(* IEC 61131-3 sources: plc-st-coding-agent/progress/evidence/f14_v13_self_20261113/jobs/custom_deepseek-v4pro (part 2) *)

(* ---- public-hard-01.raw_candidate_02.st ---- *)
(*
ENGINEERING_CONTRACT
Outputs/state group | activation | retention/hold | reset/deactivation | same-scan priority | units/bounds
estop: highest priority; active-low; all outputs false and internal states/latches reset (PUB001, PUB003).
Manual valve/motor: rising button toggles local latch; held between scans; reset by estop or mode change (PUB002, PUB004-PUB005).
AutoState: idle all off; fillA A on until level>=50; fillB B on until level>=80; processMode false->mix, true->fillC C on until level>=100; mix motor on until complete signal false->true while motor running; deliver D on and retained until autoStart/estop/mode change (PUB006-PUB015).
AutoStart rising restarts at fillA and suppresses threshold transition for first scan; transitions update state before output mapping this scan.
levelSensor INT cm; thresholds use >=.
mix completion uses armed condition requiring mixMotorComplete FALSE before TRUE while in mix state.
*)
(* CONTRACT_RULES [] *)
FUNCTION_BLOCK MaterialProportioningControl
VAR_INPUT
    estop : BOOL;
    opeMode : BOOL;
    valveAStart : BOOL;
    valveBStart : BOOL;
    valveCStart : BOOL;
    valveDStart : BOOL;
    mixMotorStart : BOOL;
    autoStart : BOOL;
    processMode : BOOL;
    levelSensor : INT;
    mixMotorComplete : BOOL;
END_VAR
VAR_OUTPUT
    valveARun : BOOL;
    valveBRun : BOOL;
    valveCRun : BOOL;
    valveDRun : BOOL;
    mixMotorRun : BOOL;
END_VAR
VAR CONSTANT
    AUTO_IDLE : INT := 0;
    AUTO_FILL_A : INT := 1;
    AUTO_FILL_B : INT := 2;
    AUTO_FILL_C : INT := 3;
    AUTO_MIX : INT := 4;
    AUTO_DELIVER : INT := 5;
END_VAR
VAR
    autoStartRtr : R_TRIG;
    valveAStartRtr : R_TRIG;
    valveBStartRtr : R_TRIG;
    valveCStartRtr : R_TRIG;
    valveDStartRtr : R_TRIG;
    mixMotorStartRtr : R_TRIG;

    local_prevOpeMode : BOOL := FALSE;
    local_init : BOOL := FALSE;

    local_manualA : BOOL := FALSE;
    local_manualB : BOOL := FALSE;
    local_manualC : BOOL := FALSE;
    local_manualD : BOOL := FALSE;
    local_manualMix : BOOL := FALSE;

    local_autoState : INT := AUTO_IDLE;
    local_firstAutoScan : BOOL := FALSE;
    local_mixArmed : BOOL := FALSE;

    local_autoStartEdge : BOOL;
    local_edgeA : BOOL;
    local_edgeB : BOOL;
    local_edgeC : BOOL;
    local_edgeD : BOOL;
    local_edgeMix : BOOL;
END_VAR

autoStartRtr(CLK := autoStart);
valveAStartRtr(CLK := valveAStart);
valveBStartRtr(CLK := valveBStart);
valveCStartRtr(CLK := valveCStart);
valveDStartRtr(CLK := valveDStart);
mixMotorStartRtr(CLK := mixMotorStart);

local_autoStartEdge := autoStartRtr.Q AND opeMode AND estop;
local_edgeA := valveAStartRtr.Q AND NOT opeMode AND estop;
local_edgeB := valveBStartRtr.Q AND NOT opeMode AND estop;
local_edgeC := valveCStartRtr.Q AND NOT opeMode AND estop;
local_edgeD := valveDStartRtr.Q AND NOT opeMode AND estop;
local_edgeMix := mixMotorStartRtr.Q AND NOT opeMode AND estop;

IF NOT local_init THEN
    local_prevOpeMode := opeMode;
    local_init := TRUE;
ELSIF local_prevOpeMode <> opeMode THEN
    local_prevOpeMode := opeMode;
    local_manualA := FALSE;
    local_manualB := FALSE;
    local_manualC := FALSE;
    local_manualD := FALSE;
    local_manualMix := FALSE;
    local_autoState := AUTO_IDLE;
    local_firstAutoScan := FALSE;
    local_mixArmed := FALSE;
END_IF;

IF NOT estop THEN
    valveARun := FALSE;
    valveBRun := FALSE;
    valveCRun := FALSE;
    valveDRun := FALSE;
    mixMotorRun := FALSE;

    local_manualA := FALSE;
    local_manualB := FALSE;
    local_manualC := FALSE;
    local_manualD := FALSE;
    local_manualMix := FALSE;
    local_autoState := AUTO_IDLE;
    local_firstAutoScan := FALSE;
    local_mixArmed := FALSE;
    RETURN;
END_IF;

IF opeMode THEN
    IF local_autoStartEdge THEN
        local_autoState := AUTO_FILL_A;
        local_firstAutoScan := TRUE;
        local_mixArmed := FALSE;
    END_IF;

    IF NOT local_firstAutoScan THEN
        IF local_autoState = AUTO_FILL_A THEN
            IF levelSensor >= 50 THEN
                local_autoState := AUTO_FILL_B;
            END_IF;
        ELSIF local_autoState = AUTO_FILL_B THEN
            IF levelSensor >= 80 THEN
                IF processMode THEN
                    local_autoState := AUTO_FILL_C;
                ELSE
                    local_autoState := AUTO_MIX;
                END_IF;
            END_IF;
        ELSIF local_autoState = AUTO_FILL_C THEN
            IF levelSensor >= 100 THEN
                local_autoState := AUTO_MIX;
            END_IF;
        ELSIF local_autoState = AUTO_MIX THEN
            IF local_mixArmed AND mixMotorComplete THEN
                local_autoState := AUTO_DELIVER;
            END_IF;
        END_IF;
    END_IF;

    IF local_autoState = AUTO_MIX THEN
        IF NOT mixMotorComplete THEN
            local_mixArmed := TRUE;
        END_IF;
    ELSE
        local_mixArmed := FALSE;
    END_IF;

    CASE local_autoState OF
        AUTO_IDLE:
            valveARun := FALSE;
            valveBRun := FALSE;
            valveCRun := FALSE;
            valveDRun := FALSE;
            mixMotorRun := FALSE;

        AUTO_FILL_A:
            valveARun := TRUE;
            valveBRun := FALSE;
            valveCRun := FALSE;
            valveDRun := FALSE;
            mixMotorRun := FALSE;

        AUTO_FILL_B:
            valveARun := FALSE;
            valveBRun := TRUE;
            valveCRun := FALSE;
            valveDRun := FALSE;
            mixMotorRun := FALSE;

        AUTO_FILL_C:
            valveARun := FALSE;
            valveBRun := FALSE;
            valveCRun := TRUE;
            valveDRun := FALSE;
            mixMotorRun := FALSE;

        AUTO_MIX:
            valveARun := FALSE;
            valveBRun := FALSE;
            valveCRun := FALSE;
            valveDRun := FALSE;
            mixMotorRun := TRUE;

        AUTO_DELIVER:
            valveARun := FALSE;
            valveBRun := FALSE;
            valveCRun := FALSE;
            valveDRun := TRUE;
            mixMotorRun := FALSE;
    END_CASE;

    local_firstAutoScan := FALSE;
ELSE
    IF local_edgeA THEN
        local_manualA := NOT local_manualA;
    END_IF;

    IF local_edgeB THEN
        local_manualB := NOT local_manualB;
    END_IF;

    IF local_edgeC THEN
        local_manualC := NOT local_manualC;
    END_IF;

    IF local_edgeD THEN
        local_manualD := NOT local_manualD;
    END_IF;

    IF local_edgeMix THEN
        local_manualMix := NOT local_manualMix;
    END_IF;

    valveARun := local_manualA;
    valveBRun := local_manualB;
    valveCRun := local_manualC;
    valveDRun := local_manualD;
    mixMotorRun := local_manualMix;
END_IF;
END_FUNCTION_BLOCK

(* ---- public-hard-02.candidate_01.st ---- *)
(*
ENGINEERING_CONTRACT
- State machine: 0=IDLE, 1=MOVING, 2=WAIT_COMPLETE, 3=DONE.
- IDLE->MOVING on rising edge of station1Start while sensor1; loads first active entry (PUB001).
- MOVING drives conveyor direction from targetStation-currentStation; stops same scan target sensor TRUE (PUB002/PUB005).
- Arrival at stations 2..4 enters WAIT_COMPLETE; arrival at 5 enters DONE (PUB003).
- WAIT_COMPLETE waits for the matching stationXComplete rising edge, then loads next entry; final 5 ends DONE (PUB003).
- Conveyor outputs are state/direction combinational and are not retained once movement stops; opposite directions cannot overlap (PUB004, V12.1).
- No unstated reset or new-cycle restart after DONE.
- Inputs are assumed valid: processLength 1..8, entries 2..5, final 5.
*)
(* CONTRACT_RULES [] *)
FUNCTION_BLOCK FlexibleProcessingControl
VAR_INPUT
    processLength : USINT;
    sensor1 : BOOL;
    sensor2 : BOOL;
    sensor3 : BOOL;
    sensor4 : BOOL;
    sensor5 : BOOL;
    station1Start : BOOL;
    station2Complete : BOOL;
    station3Complete : BOOL;
    station4Complete : BOOL;
    processSequence : ARRAY[1..8] OF USINT;
END_VAR
VAR_OUTPUT
    conveyorLeft : BOOL;
    conveyorRight : BOOL;
END_VAR
VAR
    state : INT := 0; (* 0 IDLE, 1 MOVING, 2 WAIT_COMPLETE, 3 DONE *)
    idx : USINT := 1;
    currentStation : USINT := 1;
    targetStation : USINT := 5;
    directionRight : BOOL := TRUE;
    targetArrived : BOOL := FALSE;
    completionQ : BOOL := FALSE;
    startTrig : R_TRIG;
    comp2Trig : R_TRIG;
    comp3Trig : R_TRIG;
    comp4Trig : R_TRIG;
END_VAR

startTrig(CLK := station1Start);
comp2Trig(CLK := station2Complete);
comp3Trig(CLK := station3Complete);
comp4Trig(CLK := station4Complete);

CASE targetStation OF
    2: targetArrived := sensor2;
    3: targetArrived := sensor3;
    4: targetArrived := sensor4;
    5: targetArrived := sensor5;
ELSE
    targetArrived := FALSE;
END_CASE;

IF processLength = 0 OR processLength > 8 THEN
    state := 3;
ELSE
    CASE state OF
        0: (* IDLE *)
            IF startTrig.Q AND sensor1 THEN
                idx := 1;
                currentStation := 1;
                targetStation := processSequence[idx];
                IF targetStation >= 2 AND targetStation <= 5 THEN
                    directionRight := targetStation > currentStation;
                    CASE targetStation OF
                        2: targetArrived := sensor2;
                        3: targetArrived := sensor3;
                        4: targetArrived := sensor4;
                        5: targetArrived := sensor5;
                    END_CASE;
                    IF targetArrived THEN
                        currentStation := targetStation;
                        IF targetStation = 5 THEN
                            state := 3;
                        ELSE
                            state := 2;
                        END_IF;
                    ELSE
                        state := 1;
                    END_IF;
                ELSE
                    state := 3;
                END_IF;
            END_IF;

        1: (* MOVING *)
            IF targetArrived THEN
                currentStation := targetStation;
                IF targetStation = 5 THEN
                    state := 3;
                ELSE
                    state := 2;
                END_IF;
            END_IF;

        2: (* WAIT_COMPLETE *)
            completionQ := FALSE;
            CASE currentStation OF
                2: completionQ := comp2Trig.Q;
                3: completionQ := comp3Trig.Q;
                4: completionQ := comp4Trig.Q;
            ELSE
                state := 3;
            END_CASE;
            IF completionQ THEN
                idx := idx + 1;
                IF idx > processLength THEN
                    state := 3;
                ELSE
                    targetStation := processSequence[idx];
                    IF targetStation >= 2 AND targetStation <= 5 THEN
                        directionRight := targetStation > currentStation;
                        CASE targetStation OF
                            2: targetArrived := sensor2;
                            3: targetArrived := sensor3;
                            4: targetArrived := sensor4;
                            5: targetArrived := sensor5;
                        END_CASE;
                        IF targetArrived THEN
                            currentStation := targetStation;
                            IF targetStation = 5 THEN
                                state := 3;
                            ELSE
                                state := 2;
                            END_IF;
                        ELSE
                            state := 1;
                        END_IF;
                    ELSE
                        state := 3;
                    END_IF;
                END_IF;
            END_IF;

        3: (* DONE *)
            (* no action *)
    END_CASE;
END_IF;

IF state = 1 THEN
    IF directionRight THEN
        conveyorRight := TRUE;
        conveyorLeft := FALSE;
    ELSE
        conveyorLeft := TRUE;
        conveyorRight := FALSE;
    END_IF;
ELSE
    conveyorLeft := FALSE;
    conveyorRight := FALSE;
END_IF;

END_FUNCTION_BLOCK

(* ---- public-hard-02.candidate_03.st ---- *)
(*
ENGINEERING_CONTRACT
- State machine: 0=IDLE, 1=MOVING, 2=WAIT_COMPLETE, 3=DONE.
- IDLE->MOVING on rising edge of station1Start while sensor1; loads first active entry (PUB001).
- MOVING drives conveyor direction from targetStation-currentStation; stops same scan target sensor TRUE (PUB002/PUB005).
- Arrival at stations 2..4 enters WAIT_COMPLETE; arrival at 5 enters DONE (PUB003).
- WAIT_COMPLETE waits for the matching stationXComplete rising edge, then loads next entry; final 5 ends DONE (PUB003).
- Conveyor outputs are state/direction combinational and are not retained once movement stops; opposite directions cannot overlap (PUB004, V12.1).
- No unstated reset or new-cycle restart after DONE.
- Inputs are assumed valid: processLength 1..8, entries 2..5, final 5.
*)
(* CONTRACT_RULES [] *)
FUNCTION_BLOCK FlexibleProcessingControl
VAR_INPUT
    processLength : USINT;
    sensor1 : BOOL;
    sensor2 : BOOL;
    sensor3 : BOOL;
    sensor4 : BOOL;
    sensor5 : BOOL;
    station1Start : BOOL;
    station2Complete : BOOL;
    station3Complete : BOOL;
    station4Complete : BOOL;
    processSequence : ARRAY[1..8] OF USINT;
END_VAR
VAR_OUTPUT
    conveyorLeft : BOOL;
    conveyorRight : BOOL;
END_VAR
VAR
    state : INT := 0; (* 0 IDLE, 1 MOVING, 2 WAIT_COMPLETE, 3 DONE *)
    idx : USINT := 1;
    currentStation : USINT := 1;
    targetStation : USINT := 5;
    directionRight : BOOL := TRUE;
    targetArrived : BOOL := FALSE;
    completionQ : BOOL := FALSE;
    startTrig : R_TRIG;
    comp2Trig : R_TRIG;
    comp3Trig : R_TRIG;
    comp4Trig : R_TRIG;
END_VAR

startTrig(CLK := station1Start);
comp2Trig(CLK := station2Complete);
comp3Trig(CLK := station3Complete);
comp4Trig(CLK := station4Complete);

CASE targetStation OF
    2: targetArrived := sensor2;
    3: targetArrived := sensor3;
    4: targetArrived := sensor4;
    5: targetArrived := sensor5;
ELSE
    targetArrived := FALSE;
END_CASE;

IF processLength = 0 OR processLength > 8 THEN
    state := 3;
ELSE
    CASE state OF
        0: (* IDLE *)
            IF startTrig.Q AND sensor1 THEN
                idx := 1;
                currentStation := 1;
                targetStation := processSequence[idx];
                IF targetStation >= 2 AND targetStation <= 5 THEN
                    directionRight := targetStation > currentStation;
                    CASE targetStation OF
                        2: targetArrived := sensor2;
                        3: targetArrived := sensor3;
                        4: targetArrived := sensor4;
                        5: targetArrived := sensor5;
                    END_CASE;
                    IF targetArrived THEN
                        currentStation := targetStation;
                        IF targetStation = 5 THEN
                            state := 3;
                        ELSE
                            state := 2;
                        END_IF;
                    ELSE
                        state := 1;
                    END_IF;
                ELSE
                    state := 3;
                END_IF;
            END_IF;

        1: (* MOVING *)
            IF targetArrived THEN
                currentStation := targetStation;
                IF targetStation = 5 THEN
                    state := 3;
                ELSE
                    state := 2;
                END_IF;
            END_IF;

        2: (* WAIT_COMPLETE *)
            completionQ := FALSE;
            CASE currentStation OF
                2: completionQ := comp2Trig.Q;
                3: completionQ := comp3Trig.Q;
                4: completionQ := comp4Trig.Q;
            ELSE
                state := 3;
            END_CASE;
            IF completionQ THEN
                idx := idx + 1;
                IF idx > processLength THEN
                    state := 3;
                ELSE
                    targetStation := processSequence[idx];
                    IF targetStation >= 2 AND targetStation <= 5 THEN
                        IF targetStation = currentStation THEN
                            targetArrived := TRUE;
                        ELSE
                            directionRight := targetStation > currentStation;
                            CASE targetStation OF
                                2: targetArrived := sensor2;
                                3: targetArrived := sensor3;
                                4: targetArrived := sensor4;
                                5: targetArrived := sensor5;
                            END_CASE;
                        END_IF;
                        IF targetArrived THEN
                            currentStation := targetStation;
                            IF targetStation = 5 THEN
                                state := 3;
                            ELSE
                                state := 2;
                            END_IF;
                        ELSE
                            state := 1;
                        END_IF;
                    ELSE
                        state := 3;
                    END_IF;
                END_IF;
            END_IF;

        3: (* DONE *)
            state := 0;
    END_CASE;
END_IF;

IF state = 1 THEN
    IF directionRight THEN
        conveyorRight := TRUE;
        conveyorLeft := FALSE;
    ELSE
        conveyorLeft := TRUE;
        conveyorRight := FALSE;
    END_IF;
ELSE
    conveyorLeft := FALSE;
    conveyorRight := FALSE;
END_IF;

END_FUNCTION_BLOCK

(* ---- public-hard-02.patch_base_02.st ---- *)
(*
ENGINEERING_CONTRACT
- State machine: 0=IDLE, 1=MOVING, 2=WAIT_COMPLETE, 3=DONE.
- IDLE->MOVING on rising edge of station1Start while sensor1; loads first active entry (PUB001).
- MOVING drives conveyor direction from targetStation-currentStation; stops same scan target sensor TRUE (PUB002/PUB005).
- Arrival at stations 2..4 enters WAIT_COMPLETE; arrival at 5 enters DONE (PUB003).
- WAIT_COMPLETE waits for the matching stationXComplete rising edge, then loads next entry; final 5 ends DONE (PUB003).
- Conveyor outputs are state/direction combinational and are not retained once movement stops; opposite directions cannot overlap (PUB004, V12.1).
- No unstated reset or new-cycle restart after DONE.
- Inputs are assumed valid: processLength 1..8, entries 2..5, final 5.
*)
(* CONTRACT_RULES [] *)
FUNCTION_BLOCK FlexibleProcessingControl
VAR_INPUT
    processLength : USINT;
    sensor1 : BOOL;
    sensor2 : BOOL;
    sensor3 : BOOL;
    sensor4 : BOOL;
    sensor5 : BOOL;
    station1Start : BOOL;
    station2Complete : BOOL;
    station3Complete : BOOL;
    station4Complete : BOOL;
    processSequence : ARRAY[1..8] OF USINT;
END_VAR
VAR_OUTPUT
    conveyorLeft : BOOL;
    conveyorRight : BOOL;
END_VAR
VAR
    state : INT := 0; (* 0 IDLE, 1 MOVING, 2 WAIT_COMPLETE, 3 DONE *)
    idx : USINT := 1;
    currentStation : USINT := 1;
    targetStation : USINT := 5;
    directionRight : BOOL := TRUE;
    targetArrived : BOOL := FALSE;
    completionQ : BOOL := FALSE;
    startTrig : R_TRIG;
    comp2Trig : R_TRIG;
    comp3Trig : R_TRIG;
    comp4Trig : R_TRIG;
END_VAR

startTrig(CLK := station1Start);
comp2Trig(CLK := station2Complete);
comp3Trig(CLK := station3Complete);
comp4Trig(CLK := station4Complete);

CASE targetStation OF
    2: targetArrived := sensor2;
    3: targetArrived := sensor3;
    4: targetArrived := sensor4;
    5: targetArrived := sensor5;
ELSE
    targetArrived := FALSE;
END_CASE;

IF processLength = 0 OR processLength > 8 THEN
    state := 3;
ELSE
    CASE state OF
        0: (* IDLE *)
            IF startTrig.Q AND sensor1 THEN
                idx := 1;
                currentStation := 1;
                targetStation := processSequence[idx];
                IF targetStation >= 2 AND targetStation <= 5 THEN
                    directionRight := targetStation > currentStation;
                    CASE targetStation OF
                        2: targetArrived := sensor2;
                        3: targetArrived := sensor3;
                        4: targetArrived := sensor4;
                        5: targetArrived := sensor5;
                    END_CASE;
                    IF targetArrived THEN
                        currentStation := targetStation;
                        IF targetStation = 5 THEN
                            state := 3;
                        ELSE
                            state := 2;
                        END_IF;
                    ELSE
                        state := 1;
                    END_IF;
                ELSE
                    state := 3;
                END_IF;
            END_IF;

        1: (* MOVING *)
            IF targetArrived THEN
                currentStation := targetStation;
                IF targetStation = 5 THEN
                    state := 3;
                ELSE
                    state := 2;
                END_IF;
            END_IF;

        2: (* WAIT_COMPLETE *)
            completionQ := FALSE;
            CASE currentStation OF
                2: completionQ := comp2Trig.Q;
                3: completionQ := comp3Trig.Q;
                4: completionQ := comp4Trig.Q;
            ELSE
                state := 3;
            END_CASE;
            IF completionQ THEN
                idx := idx + 1;
                IF idx > processLength THEN
                    state := 3;
                ELSE
                    targetStation := processSequence[idx];
                    IF targetStation >= 2 AND targetStation <= 5 THEN
                        directionRight := targetStation > currentStation;
                        CASE targetStation OF
                            2: targetArrived := sensor2;
                            3: targetArrived := sensor3;
                            4: targetArrived := sensor4;
                            5: targetArrived := sensor5;
                        END_CASE;
                        IF targetArrived THEN
                            currentStation := targetStation;
                            IF targetStation = 5 THEN
                                state := 3;
                            ELSE
                                state := 2;
                            END_IF;
                        ELSE
                            state := 1;
                        END_IF;
                    ELSE
                        state := 3;
                    END_IF;
                END_IF;
            END_IF;

        3: (* DONE *)
            (* no action *)
    END_CASE;
END_IF;

IF state = 1 THEN
    IF directionRight THEN
        conveyorRight := TRUE;
        conveyorLeft := FALSE;
    ELSE
        conveyorLeft := TRUE;
        conveyorRight := FALSE;
    END_IF;
ELSE
    conveyorLeft := FALSE;
    conveyorRight := FALSE;
END_IF;

END_FUNCTION_BLOCK

(* ---- public-hard-02.patch_base_03.st ---- *)
(*
ENGINEERING_CONTRACT
- State machine: 0=IDLE, 1=MOVING, 2=WAIT_COMPLETE, 3=DONE.
- IDLE->MOVING on rising edge of station1Start while sensor1; loads first active entry (PUB001).
- MOVING drives conveyor direction from targetStation-currentStation; stops same scan target sensor TRUE (PUB002/PUB005).
- Arrival at stations 2..4 enters WAIT_COMPLETE; arrival at 5 enters DONE (PUB003).
- WAIT_COMPLETE waits for the matching stationXComplete rising edge, then loads next entry; final 5 ends DONE (PUB003).
- Conveyor outputs are state/direction combinational and are not retained once movement stops; opposite directions cannot overlap (PUB004, V12.1).
- No unstated reset or new-cycle restart after DONE.
- Inputs are assumed valid: processLength 1..8, entries 2..5, final 5.
*)
(* CONTRACT_RULES [] *)
FUNCTION_BLOCK FlexibleProcessingControl
VAR_INPUT
    processLength : USINT;
    sensor1 : BOOL;
    sensor2 : BOOL;
    sensor3 : BOOL;
    sensor4 : BOOL;
    sensor5 : BOOL;
    station1Start : BOOL;
    station2Complete : BOOL;
    station3Complete : BOOL;
    station4Complete : BOOL;
    processSequence : ARRAY[1..8] OF USINT;
END_VAR
VAR_OUTPUT
    conveyorLeft : BOOL;
    conveyorRight : BOOL;
END_VAR
VAR
    state : INT := 0; (* 0 IDLE, 1 MOVING, 2 WAIT_COMPLETE, 3 DONE *)
    idx : USINT := 1;
    currentStation : USINT := 1;
    targetStation : USINT := 5;
    directionRight : BOOL := TRUE;
    targetArrived : BOOL := FALSE;
    completionQ : BOOL := FALSE;
    startTrig : R_TRIG;
    comp2Trig : R_TRIG;
    comp3Trig : R_TRIG;
    comp4Trig : R_TRIG;
END_VAR

startTrig(CLK := station1Start);
comp2Trig(CLK := station2Complete);
comp3Trig(CLK := station3Complete);
comp4Trig(CLK := station4Complete);

CASE targetStation OF
    2: targetArrived := sensor2;
    3: targetArrived := sensor3;
    4: targetArrived := sensor4;
    5: targetArrived := sensor5;
ELSE
    targetArrived := FALSE;
END_CASE;

IF processLength = 0 OR processLength > 8 THEN
    state := 3;
ELSE
    CASE state OF
        0: (* IDLE *)
            IF startTrig.Q AND sensor1 THEN
                idx := 1;
                currentStation := 1;
                targetStation := processSequence[idx];
                IF targetStation >= 2 AND targetStation <= 5 THEN
                    directionRight := targetStation > currentStation;
                    CASE targetStation OF
                        2: targetArrived := sensor2;
                        3: targetArrived := sensor3;
                        4: targetArrived := sensor4;
                        5: targetArrived := sensor5;
                    END_CASE;
                    IF targetArrived THEN
                        currentStation := targetStation;
                        IF targetStation = 5 THEN
                            state := 3;
                        ELSE
                            state := 2;
                        END_IF;
                    ELSE
                        state := 1;
                    END_IF;
                ELSE
                    state := 3;
                END_IF;
            END_IF;

        1: (* MOVING *)
            IF targetArrived THEN
                currentStation := targetStation;
                IF targetStation = 5 THEN
                    state := 3;
                ELSE
                    state := 2;
                END_IF;
            END_IF;

        2: (* WAIT_COMPLETE *)
            completionQ := FALSE;
            CASE currentStation OF
                2: completionQ := comp2Trig.Q;
                3: completionQ := comp3Trig.Q;
                4: completionQ := comp4Trig.Q;
            ELSE
                state := 3;
            END_CASE;
            IF completionQ THEN
                idx := idx + 1;
                IF idx > processLength THEN
                    state := 3;
                ELSE
                    targetStation := processSequence[idx];
                    IF targetStation >= 2 AND targetStation <= 5 THEN
                        directionRight := targetStation > currentStation;
                        CASE targetStation OF
                            2: targetArrived := sensor2;
                            3: targetArrived := sensor3;
                            4: targetArrived := sensor4;
                            5: targetArrived := sensor5;
                        END_CASE;
                        IF targetArrived THEN
                            currentStation := targetStation;
                            IF targetStation = 5 THEN
                                state := 3;
                            ELSE
                                state := 2;
                            END_IF;
                        ELSE
                            state := 1;
                        END_IF;
                    ELSE
                        state := 3;
                    END_IF;
                END_IF;
            END_IF;

        3: (* DONE *)
            (* no action *)
    END_CASE;
END_IF;

IF state = 1 THEN
    IF directionRight THEN
        conveyorRight := TRUE;
        conveyorLeft := FALSE;
    ELSE
        conveyorLeft := TRUE;
        conveyorRight := FALSE;
    END_IF;
ELSE
    conveyorLeft := FALSE;
    conveyorRight := FALSE;
END_IF;

END_FUNCTION_BLOCK

(* ---- public-hard-02.raw_candidate_01.st ---- *)
(*
ENGINEERING_CONTRACT
- State machine: 0=IDLE, 1=MOVING, 2=WAIT_COMPLETE, 3=DONE.
- IDLE->MOVING on rising edge of station1Start while sensor1; loads first active entry (PUB001).
- MOVING drives conveyor direction from targetStation-currentStation; stops same scan target sensor TRUE (PUB002/PUB005).
- Arrival at stations 2..4 enters WAIT_COMPLETE; arrival at 5 enters DONE (PUB003).
- WAIT_COMPLETE waits for the matching stationXComplete rising edge, then loads next entry; final 5 ends DONE (PUB003).
- Conveyor outputs are state/direction combinational and are not retained once movement stops; opposite directions cannot overlap (PUB004, V12.1).
- No unstated reset or new-cycle restart after DONE.
- Inputs are assumed valid: processLength 1..8, entries 2..5, final 5.
*)
(* CONTRACT_RULES [] *)
FUNCTION_BLOCK FlexibleProcessingControl
VAR_INPUT
    processLength : USINT;
    sensor1 : BOOL;
    sensor2 : BOOL;
    sensor3 : BOOL;
    sensor4 : BOOL;
    sensor5 : BOOL;
    station1Start : BOOL;
    station2Complete : BOOL;
    station3Complete : BOOL;
    station4Complete : BOOL;
    processSequence : ARRAY[1..8] OF USINT;
END_VAR
VAR_OUTPUT
    conveyorLeft : BOOL;
    conveyorRight : BOOL;
END_VAR
VAR
    state : INT := 0; (* 0 IDLE, 1 MOVING, 2 WAIT_COMPLETE, 3 DONE *)
    idx : USINT := 1;
    currentStation : USINT := 1;
    targetStation : USINT := 5;
    directionRight : BOOL := TRUE;
    targetArrived : BOOL := FALSE;
    completionQ : BOOL := FALSE;
    startTrig : R_TRIG;
    comp2Trig : R_TRIG;
    comp3Trig : R_TRIG;
    comp4Trig : R_TRIG;
END_VAR

startTrig(CLK := station1Start);
comp2Trig(CLK := station2Complete);
comp3Trig(CLK := station3Complete);
comp4Trig(CLK := station4Complete);

CASE targetStation OF
    2: targetArrived := sensor2;
    3: targetArrived := sensor3;
    4: targetArrived := sensor4;
    5: targetArrived := sensor5;
ELSE
    targetArrived := FALSE;
END_CASE

IF processLength = 0 OR processLength > 8 THEN
    state := 3;
ELSE
    CASE state OF
        0: (* IDLE *)
            IF startTrig.Q AND sensor1 THEN
                idx := 1;
                currentStation := 1;
                targetStation := processSequence[idx];
                IF targetStation >= 2 AND targetStation <= 5 THEN
                    directionRight := targetStation > currentStation;
                    CASE targetStation OF
                        2: targetArrived := sensor2;
                        3: targetArrived := sensor3;
                        4: targetArrived := sensor4;
                        5: targetArrived := sensor5;
                    END_CASE
                    IF targetArrived THEN
                        currentStation := targetStation;
                        IF targetStation = 5 THEN
                            state := 3;
                        ELSE
                            state := 2;
                        END_IF
                    ELSE
                        state := 1;
                    END_IF
                ELSE
                    state := 3;
                END_IF
            END_IF

        1: (* MOVING *)
            IF targetArrived THEN
                currentStation := targetStation;
                IF targetStation = 5 THEN
                    state := 3;
                ELSE
                    state := 2;
                END_IF
            END_IF

        2: (* WAIT_COMPLETE *)
            completionQ := FALSE;
            CASE currentStation OF
                2: completionQ := comp2Trig.Q;
                3: completionQ := comp3Trig.Q;
                4: completionQ := comp4Trig.Q;
            ELSE
                state := 3;
            END_CASE
            IF completionQ THEN
                idx := idx + 1;
                IF idx > processLength THEN
                    state := 3;
                ELSE
                    targetStation := processSequence[idx];
                    IF targetStation >= 2 AND targetStation <= 5 THEN
                        directionRight := targetStation > currentStation;
                        CASE targetStation OF
                            2: targetArrived := sensor2;
                            3: targetArrived := sensor3;
                            4: targetArrived := sensor4;
                            5: targetArrived := sensor5;
                        END_CASE
                        IF targetArrived THEN
                            currentStation := targetStation;
                            IF targetStation = 5 THEN
                                state := 3;
                            ELSE
                                state := 2;
                            END_IF
                        ELSE
                            state := 1;
                        END_IF
                    ELSE
                        state := 3;
                    END_IF
                END_IF
            END_IF

        3: (* DONE *)
            (* no action *)
    END_CASE
END_IF

IF state = 1 THEN
    IF directionRight THEN
        conveyorRight := TRUE;
        conveyorLeft := FALSE;
    ELSE
        conveyorLeft := TRUE;
        conveyorRight := FALSE;
    END_IF
ELSE
    conveyorLeft := FALSE;
    conveyorRight := FALSE;
END_IF

END_FUNCTION_BLOCK

(* ---- public-hard-02.raw_candidate_03.st ---- *)
(*
ENGINEERING_CONTRACT
- State machine: 0=IDLE, 1=MOVING, 2=WAIT_COMPLETE, 3=DONE.
- IDLE->MOVING on rising edge of station1Start while sensor1; loads first active entry (PUB001).
- MOVING drives conveyor direction from targetStation-currentStation; stops same scan target sensor TRUE (PUB002/PUB005).
- Arrival at stations 2..4 enters WAIT_COMPLETE; arrival at 5 enters DONE (PUB003).
- WAIT_COMPLETE waits for the matching stationXComplete rising edge, then loads next entry; final 5 ends DONE (PUB003).
- Conveyor outputs are state/direction combinational and are not retained once movement stops; opposite directions cannot overlap (PUB004, V12.1).
- No unstated reset or new-cycle restart after DONE.
- Inputs are assumed valid: processLength 1..8, entries 2..5, final 5.
*)
(* CONTRACT_RULES [] *)
FUNCTION_BLOCK FlexibleProcessingControl
VAR_INPUT
    processLength : USINT;
    sensor1 : BOOL;
    sensor2 : BOOL;
    sensor3 : BOOL;
    sensor4 : BOOL;
    sensor5 : BOOL;
    station1Start : BOOL;
    station2Complete : BOOL;
    station3Complete : BOOL;
    station4Complete : BOOL;
    processSequence : ARRAY[1..8] OF USINT;
END_VAR
VAR_OUTPUT
    conveyorLeft : BOOL;
    conveyorRight : BOOL;
END_VAR
VAR
    state : INT := 0; (* 0 IDLE, 1 MOVING, 2 WAIT_COMPLETE, 3 DONE *)
    idx : USINT := 1;
    currentStation : USINT := 1;
    targetStation : USINT := 5;
    directionRight : BOOL := TRUE;
    targetArrived : BOOL := FALSE;
    completionQ : BOOL := FALSE;
    startTrig : R_TRIG;
    comp2Trig : R_TRIG;
    comp3Trig : R_TRIG;
    comp4Trig : R_TRIG;
END_VAR

startTrig(CLK := station1Start);
comp2Trig(CLK := station2Complete);
comp3Trig(CLK := station3Complete);
comp4Trig(CLK := station4Complete);

CASE targetStation OF
    2: targetArrived := sensor2;
    3: targetArrived := sensor3;
    4: targetArrived := sensor4;
    5: targetArrived := sensor5;
ELSE
    targetArrived := FALSE;
END_CASE;

IF processLength = 0 OR processLength > 8 THEN
    state := 3;
ELSE
    CASE state OF
        0: (* IDLE *)
            IF startTrig.Q AND sensor1 THEN
                idx := 1;
                currentStation := 1;
                targetStation := processSequence[idx];
                IF targetStation >= 2 AND targetStation <= 5 THEN
                    directionRight := targetStation > currentStation;
                    CASE targetStation OF
                        2: targetArrived := sensor2;
                        3: targetArrived := sensor3;
                        4: targetArrived := sensor4;
                        5: targetArrived := sensor5;
                    END_CASE;
                    IF targetArrived THEN
                        currentStation := targetStation;
                        IF targetStation = 5 THEN
                            state := 3;
                        ELSE
                            state := 2;
                        END_IF;
                    ELSE
                        state := 1;
                    END_IF;
                ELSE
                    state := 3;
                END_IF;
            END_IF;

        1: (* MOVING *)
            IF targetArrived THEN
                currentStation := targetStation;
                IF targetStation = 5 THEN
                    state := 3;
                ELSE
                    state := 2;
                END_IF;
            END_IF;

        2: (* WAIT_COMPLETE *)
            completionQ := FALSE;
            CASE currentStation OF
                2: completionQ := comp2Trig.Q;
                3: completionQ := comp3Trig.Q;
                4: completionQ := comp4Trig.Q;
            ELSE
                state := 3;
            END_CASE;
            IF completionQ THEN
                idx := idx + 1;
                IF idx > processLength THEN
                    state := 3;
                ELSE
                    targetStation := processSequence[idx];
                    IF targetStation >= 2 AND targetStation <= 5 THEN
                        IF targetStation = currentStation THEN
                            targetArrived := TRUE;
                        ELSE
                            directionRight := targetStation > currentStation;
                            CASE targetStation OF
                                2: targetArrived := sensor2;
                                3: targetArrived := sensor3;
                                4: targetArrived := sensor4;
                                5: targetArrived := sensor5;
                            END_CASE;
                        END_IF;
                        IF targetArrived THEN
                            currentStation := targetStation;
                            IF targetStation = 5 THEN
                                state := 3;
                            ELSE
                                state := 2;
                            END_IF;
                        ELSE
                            state := 1;
                        END_IF;
                    ELSE
                        state := 3;
                    END_IF;
                END_IF;
            END_IF;

        3: (* DONE *)
            state := 0;
    END_CASE;
END_IF;

IF state = 1 THEN
    IF directionRight THEN
        conveyorRight := TRUE;
        conveyorLeft := FALSE;
    ELSE
        conveyorLeft := TRUE;
        conveyorRight := FALSE;
    END_IF;
ELSE
    conveyorLeft := FALSE;
    conveyorRight := FALSE;
END_IF;

END_FUNCTION_BLOCK

(* ---- public-hard-03.candidate_01.st ---- *)
(*
ENGINEERING_CONTRACT
- recipeAdded/Deleted/Modified: rising-edge pulse outputs, TRUE only on the scan where the corresponding request succeeds; no retention; reset next scan (PUB003/004/005).
- error: rising-edge pulse, TRUE only on the scan where an operation fails; no retention; reset next scan (PUB002-005).
- status: WORD code, 0 by default, nonzero only during a failed operation scan (PUB002-005).
- recipeQueryResult: zero-cleared at the start of every scan; holds the full recipe only during a successful query scan (PUB002).
- recipe database: persistent through IN_OUT; add uses smallest empty slot, duplicate check; delete sets recipeID to 0; modify replaces the whole struct (PUB003/004/005).
- Simultaneous requests are processed in the order query, add, delete, modify; unspecified by PUB002-005.
- recipeID 0 is treated as nonexistent for query/delete/modify and as duplicate for add because 0 marks an empty slot (PUB001).
*)
(* CONTRACT_RULES [] *)
FUNCTION_BLOCK FB_RecipeManagement
VAR_INPUT
    addRecipe : BOOL;
    deleteRecipe : BOOL;
    modifyRecipe : BOOL;
    queryRecipe : BOOL;
    recipeIn : ST_Recipe;
END_VAR

VAR_OUTPUT
    recipeAdded : BOOL;
    recipeDeleted : BOOL;
    recipeModified : BOOL;
    recipeQueryResult : ST_Recipe;
    error : BOOL;
    status : WORD;
END_VAR

VAR_IN_OUT
    recipe : ARRAY[1..10] OF ST_Recipe;
END_VAR

VAR
    tmp_TrigAdd : R_TRIG;
    tmp_TrigDelete : R_TRIG;
    tmp_TrigModify : R_TRIG;
    tmp_TrigQuery : R_TRIG;
    tmp_idx : INT;
    tmp_found : BOOL;
    tmp_foundIdx : INT;
    tmp_emptyIdx : INT;
END_VAR

// Evaluate rising edges once per scan.
tmp_TrigAdd(CLK := addRecipe);
tmp_TrigDelete(CLK := deleteRecipe);
tmp_TrigModify(CLK := modifyRecipe);
tmp_TrigQuery(CLK := queryRecipe);

// Default outputs for this scan.
recipeAdded := FALSE;
recipeDeleted := FALSE;
recipeModified := FALSE;
error := FALSE;
status := 0;

// Clear query result each scan; successful query will overwrite later.
recipeQueryResult.recipeID := 0;
recipeQueryResult.ingredientType := 0;
recipeQueryResult.ingredientRatio := 0.0;
recipeQueryResult.productionTemperature := 0.0;

// Query operation (PUB002)
IF tmp_TrigQuery.Q THEN
    tmp_foundIdx := 0;
    IF recipeIn.recipeID <> 0 THEN
        FOR tmp_idx := 1 TO 10 DO
            IF recipe[tmp_idx].recipeID = recipeIn.recipeID THEN
                tmp_foundIdx := tmp_idx;
                EXIT;
            END_IF;
        END_FOR;
    END_IF;

    IF tmp_foundIdx = 0 THEN
        error := TRUE;
        status := 16#8001;
    ELSE
        recipeQueryResult := recipe[tmp_foundIdx];
    END_IF;
END_IF;

// Add operation (PUB003)
IF tmp_TrigAdd.Q THEN
    tmp_found := FALSE;
    tmp_emptyIdx := 0;

    FOR tmp_idx := 1 TO 10 DO
        IF recipe[tmp_idx].recipeID = recipeIn.recipeID THEN
            tmp_found := TRUE;
            EXIT;
        END_IF;
        IF recipe[tmp_idx].recipeID = 0 AND tmp_emptyIdx = 0 THEN
            tmp_emptyIdx := tmp_idx;
        END_IF;
    END_FOR;

    IF tmp_found THEN
        error := TRUE;
        status := 16#8002;
    ELSIF tmp_emptyIdx = 0 THEN
        error := TRUE;
        status := 16#8003;
    ELSE
        recipe[tmp_emptyIdx] := recipeIn;
        recipeAdded := TRUE;
    END_IF;
END_IF;

// Delete operation (PUB004)
IF tmp_TrigDelete.Q THEN
    tmp_foundIdx := 0;
    IF recipeIn.recipeID <> 0 THEN
        FOR tmp_idx := 1 TO 10 DO
            IF recipe[tmp_idx].recipeID = recipeIn.recipeID THEN
                tmp_foundIdx := tmp_idx;
                EXIT;
            END_IF;
        END_FOR;
    END_IF;

    IF tmp_foundIdx = 0 THEN
        error := TRUE;
        status := 16#8004;
    ELSE
        recipe[tmp_foundIdx].recipeID := 0;
        recipeDeleted := TRUE;
    END_IF;
END_IF;

// Modify operation (PUB005)
IF tmp_TrigModify.Q THEN
    tmp_foundIdx := 0;
    IF recipeIn.recipeID <> 0 THEN
        FOR tmp_idx := 1 TO 10 DO
            IF recipe[tmp_idx].recipeID = recipeIn.recipeID THEN
                tmp_foundIdx := tmp_idx;
                EXIT;
            END_IF;
        END_FOR;
    END_IF;

    IF tmp_foundIdx = 0 THEN
        error := TRUE;
        status := 16#8005;
    ELSE
        recipe[tmp_foundIdx] := recipeIn;
        recipeModified := TRUE;
    END_IF;
END_IF;

END_FUNCTION_BLOCK

(* ---- public-hard-03.candidate_02.st ---- *)
(*
ENGINEERING_CONTRACT
- recipeAdded/Deleted/Modified: rising-edge pulse outputs, TRUE only on the scan where the corresponding request succeeds; no retention; reset next scan (PUB003/004/005).
- error: rising-edge pulse, TRUE only on the scan where an operation fails; no retention; reset next scan (PUB002-005).
- status: WORD code, 0 by default, nonzero only during a failed operation scan (PUB002-005).
- recipeQueryResult: zero-cleared at the start of every scan; holds the full recipe only during a successful query scan (PUB002).
- recipe database: persistent through IN_OUT; add uses smallest empty slot, duplicate check; delete sets recipeID to 0; modify replaces the whole struct (PUB003/004/005).
- Simultaneous requests are processed in the order query, add, delete, modify; unspecified by PUB002-005.
- recipeID 0 is treated as nonexistent for query/delete/modify and as duplicate for add because 0 marks an empty slot (PUB001).
*)
(* CONTRACT_RULES [] *)
TYPE ST_Recipe :
STRUCT
    recipeID : INT;
    ingredientType : INT;
    ingredientRatio : REAL;
    productionTemperature : REAL;
END_STRUCT
END_TYPE;

FUNCTION_BLOCK FB_RecipeManagement
VAR_INPUT
    addRecipe : BOOL;
    deleteRecipe : BOOL;
    modifyRecipe : BOOL;
    queryRecipe : BOOL;
    recipeIn : ST_Recipe;
END_VAR

VAR_OUTPUT
    recipeAdded : BOOL;
    recipeDeleted : BOOL;
    recipeModified : BOOL;
    recipeQueryResult : ST_Recipe;
    error : BOOL;
    status : WORD;
END_VAR

VAR_IN_OUT
    recipe : ARRAY[1..10] OF ST_Recipe;
END_VAR

VAR
    tmp_TrigAdd : R_TRIG;
    tmp_TrigDelete : R_TRIG;
    tmp_TrigModify : R_TRIG;
    tmp_TrigQuery : R_TRIG;
    tmp_idx : INT;
    tmp_found : BOOL;
    tmp_foundIdx : INT;
    tmp_emptyIdx : INT;
END_VAR

// Evaluate rising edges once per scan.
tmp_TrigAdd(CLK := addRecipe);
tmp_TrigDelete(CLK := deleteRecipe);
tmp_TrigModify(CLK := modifyRecipe);
tmp_TrigQuery(CLK := queryRecipe);

// Default outputs for this scan.
recipeAdded := FALSE;
recipeDeleted := FALSE;
recipeModified := FALSE;
error := FALSE;
status := 0;

// Clear query result each scan; successful query will overwrite later.
recipeQueryResult.recipeID := 0;
recipeQueryResult.ingredientType := 0;
recipeQueryResult.ingredientRatio := 0.0;
recipeQueryResult.productionTemperature := 0.0;

// Query operation (PUB002)
IF tmp_TrigQuery.Q THEN
    tmp_foundIdx := 0;
    IF recipeIn.recipeID <> 0 THEN
        FOR tmp_idx := 1 TO 10 DO
            IF recipe[tmp_idx].recipeID = recipeIn.recipeID THEN
                tmp_foundIdx := tmp_idx;
                EXIT;
            END_IF;
        END_FOR;
    END_IF;

    IF tmp_foundIdx = 0 THEN
        error := TRUE;
        status := 16#8001;
    ELSE
        recipeQueryResult := recipe[tmp_foundIdx];
    END_IF;
END_IF;

// Add operation (PUB003)
IF tmp_TrigAdd.Q THEN
    tmp_found := FALSE;
    tmp_emptyIdx := 0;

    FOR tmp_idx := 1 TO 10 DO
        IF recipe[tmp_idx].recipeID = recipeIn.recipeID THEN
            tmp_found := TRUE;
            EXIT;
        END_IF;
        IF recipe[tmp_idx].recipeID = 0 AND tmp_emptyIdx = 0 THEN
            tmp_emptyIdx := tmp_idx;
        END_IF;
    END_FOR;

    IF tmp_found THEN
        error := TRUE;
        status := 16#8002;
    ELSIF tmp_emptyIdx = 0 THEN
        error := TRUE;
        status := 16#8003;
    ELSE
        recipe[tmp_emptyIdx] := recipeIn;
        recipeAdded := TRUE;
    END_IF;
END_IF;

// Delete operation (PUB004)
IF tmp_TrigDelete.Q THEN
    tmp_foundIdx := 0;
    IF recipeIn.recipeID <> 0 THEN
        FOR tmp_idx := 1 TO 10 DO
            IF recipe[tmp_idx].recipeID = recipeIn.recipeID THEN
                tmp_foundIdx := tmp_idx;
                EXIT;
            END_IF;
        END_FOR;
    END_IF;

    IF tmp_foundIdx = 0 THEN
        error := TRUE;
        status := 16#8004;
    ELSE
        recipe[tmp_foundIdx].recipeID := 0;
        recipeDeleted := TRUE;
    END_IF;
END_IF;

// Modify operation (PUB005)
IF tmp_TrigModify.Q THEN
    tmp_foundIdx := 0;
    IF recipeIn.recipeID <> 0 THEN
        FOR tmp_idx := 1 TO 10 DO
            IF recipe[tmp_idx].recipeID = recipeIn.recipeID THEN
                tmp_foundIdx := tmp_idx;
                EXIT;
            END_IF;
        END_FOR;
    END_IF;

    IF tmp_foundIdx = 0 THEN
        error := TRUE;
        status := 16#8005;
    ELSE
        recipe[tmp_foundIdx] := recipeIn;
        recipeModified := TRUE;
    END_IF;
END_IF;

END_FUNCTION_BLOCK

(* ---- public-hard-03.patch_base_02.st ---- *)
(*
ENGINEERING_CONTRACT
- recipeAdded/Deleted/Modified: rising-edge pulse outputs, TRUE only on the scan where the corresponding request succeeds; no retention; reset next scan (PUB003/004/005).
- error: rising-edge pulse, TRUE only on the scan where an operation fails; no retention; reset next scan (PUB002-005).
- status: WORD code, 0 by default, nonzero only during a failed operation scan (PUB002-005).
- recipeQueryResult: zero-cleared at the start of every scan; holds the full recipe only during a successful query scan (PUB002).
- recipe database: persistent through IN_OUT; add uses smallest empty slot, duplicate check; delete sets recipeID to 0; modify replaces the whole struct (PUB003/004/005).
- Simultaneous requests are processed in the order query, add, delete, modify; unspecified by PUB002-005.
- recipeID 0 is treated as nonexistent for query/delete/modify and as duplicate for add because 0 marks an empty slot (PUB001).
*)
(* CONTRACT_RULES [] *)
FUNCTION_BLOCK FB_RecipeManagement
VAR_INPUT
    addRecipe : BOOL;
    deleteRecipe : BOOL;
    modifyRecipe : BOOL;
    queryRecipe : BOOL;
    recipeIn : ST_Recipe;
END_VAR

VAR_OUTPUT
    recipeAdded : BOOL;
    recipeDeleted : BOOL;
    recipeModified : BOOL;
    recipeQueryResult : ST_Recipe;
    error : BOOL;
    status : WORD;
END_VAR

VAR_IN_OUT
    recipe : ARRAY[1..10] OF ST_Recipe;
END_VAR

VAR
    tmp_TrigAdd : R_TRIG;
    tmp_TrigDelete : R_TRIG;
    tmp_TrigModify : R_TRIG;
    tmp_TrigQuery : R_TRIG;
    tmp_idx : INT;
    tmp_found : BOOL;
    tmp_foundIdx : INT;
    tmp_emptyIdx : INT;
END_VAR

// Evaluate rising edges once per scan.
tmp_TrigAdd(CLK := addRecipe);
tmp_TrigDelete(CLK := deleteRecipe);
tmp_TrigModify(CLK := modifyRecipe);
tmp_TrigQuery(CLK := queryRecipe);

// Default outputs for this scan.
recipeAdded := FALSE;
recipeDeleted := FALSE;
recipeModified := FALSE;
error := FALSE;
status := 0;

// Clear query result each scan; successful query will overwrite later.
recipeQueryResult.recipeID := 0;
recipeQueryResult.ingredientType := 0;
recipeQueryResult.ingredientRatio := 0.0;
recipeQueryResult.productionTemperature := 0.0;

// Query operation (PUB002)
IF tmp_TrigQuery.Q THEN
    tmp_foundIdx := 0;
    IF recipeIn.recipeID <> 0 THEN
        FOR tmp_idx := 1 TO 10 DO
            IF recipe[tmp_idx].recipeID = recipeIn.recipeID THEN
                tmp_foundIdx := tmp_idx;
                EXIT;
            END_IF;
        END_FOR;
    END_IF;

    IF tmp_foundIdx = 0 THEN
        error := TRUE;
        status := 16#8001;
    ELSE
        recipeQueryResult := recipe[tmp_foundIdx];
    END_IF;
END_IF;

// Add operation (PUB003)
IF tmp_TrigAdd.Q THEN
    tmp_found := FALSE;
    tmp_emptyIdx := 0;

    FOR tmp_idx := 1 TO 10 DO
        IF recipe[tmp_idx].recipeID = recipeIn.recipeID THEN
            tmp_found := TRUE;
            EXIT;
        END_IF;
        IF recipe[tmp_idx].recipeID = 0 AND tmp_emptyIdx = 0 THEN
            tmp_emptyIdx := tmp_idx;
        END_IF;
    END_FOR;

    IF tmp_found THEN
        error := TRUE;
        status := 16#8002;
    ELSIF tmp_emptyIdx = 0 THEN
        error := TRUE;
        status := 16#8003;
    ELSE
        recipe[tmp_emptyIdx] := recipeIn;
        recipeAdded := TRUE;
    END_IF;
END_IF;

// Delete operation (PUB004)
IF tmp_TrigDelete.Q THEN
    tmp_foundIdx := 0;
    IF recipeIn.recipeID <> 0 THEN
        FOR tmp_idx := 1 TO 10 DO
            IF recipe[tmp_idx].recipeID = recipeIn.recipeID THEN
                tmp_foundIdx := tmp_idx;
                EXIT;
            END_IF;
        END_FOR;
    END_IF;

    IF tmp_foundIdx = 0 THEN
        error := TRUE;
        status := 16#8004;
    ELSE
        recipe[tmp_foundIdx].recipeID := 0;
        recipeDeleted := TRUE;
    END_IF;
END_IF;

// Modify operation (PUB005)
IF tmp_TrigModify.Q THEN
    tmp_foundIdx := 0;
    IF recipeIn.recipeID <> 0 THEN
        FOR tmp_idx := 1 TO 10 DO
            IF recipe[tmp_idx].recipeID = recipeIn.recipeID THEN
                tmp_foundIdx := tmp_idx;
                EXIT;
            END_IF;
        END_FOR;
    END_IF;

    IF tmp_foundIdx = 0 THEN
        error := TRUE;
        status := 16#8005;
    ELSE
        recipe[tmp_foundIdx] := recipeIn;
        recipeModified := TRUE;
    END_IF;
END_IF;

END_FUNCTION_BLOCK

(* ---- public-hard-03.raw_candidate_01.st ---- *)
(*
ENGINEERING_CONTRACT
- recipeAdded/Deleted/Modified: rising-edge pulse outputs, TRUE only on the scan where the corresponding request succeeds; no retention; reset next scan (PUB003/004/005).
- error: rising-edge pulse, TRUE only on the scan where an operation fails; no retention; reset next scan (PUB002-005).
- status: WORD code, 0 by default, nonzero only during a failed operation scan (PUB002-005).
- recipeQueryResult: zero-cleared at the start of every scan; holds the full recipe only during a successful query scan (PUB002).
- recipe database: persistent through IN_OUT; add uses smallest empty slot, duplicate check; delete sets recipeID to 0; modify replaces the whole struct (PUB003/004/005).
- Simultaneous requests are processed in the order query, add, delete, modify; unspecified by PUB002-005.
- recipeID 0 is treated as nonexistent for query/delete/modify and as duplicate for add because 0 marks an empty slot (PUB001).
*)
(* CONTRACT_RULES [] *)
FUNCTION_BLOCK FB_RecipeManagement
VAR_INPUT
    addRecipe : BOOL;
    deleteRecipe : BOOL;
    modifyRecipe : BOOL;
    queryRecipe : BOOL;
    recipeIn : ST_Recipe;
END_VAR

VAR_OUTPUT
    recipeAdded : BOOL;
    recipeDeleted : BOOL;
    recipeModified : BOOL;
    recipeQueryResult : ST_Recipe;
    error : BOOL;
    status : WORD;
END_VAR

VAR_IN_OUT
    recipe : ARRAY[1..10] OF ST_Recipe;
END_VAR

VAR
    tmp_TrigAdd : R_TRIG;
    tmp_TrigDelete : R_TRIG;
    tmp_TrigModify : R_TRIG;
    tmp_TrigQuery : R_TRIG;
    tmp_idx : INT;
    tmp_found : BOOL;
    tmp_foundIdx : INT;
    tmp_emptyIdx : INT;
END_VAR

// Evaluate rising edges once per scan.
tmp_TrigAdd(CLK := addRecipe);
tmp_TrigDelete(CLK := deleteRecipe);
tmp_TrigModify(CLK := modifyRecipe);
tmp_TrigQuery(CLK := queryRecipe);

// Default outputs for this scan.
recipeAdded := FALSE;
recipeDeleted := FALSE;
recipeModified := FALSE;
error := FALSE;
status := 0;

// Clear query result each scan; successful query will overwrite later.
recipeQueryResult.recipeID := 0;
recipeQueryResult.ingredientType := 0;
recipeQueryResult.ingredientRatio := 0.0;
recipeQueryResult.productionTemperature := 0.0;

// Query operation (PUB002)
IF tmp_TrigQuery.Q THEN
    tmp_foundIdx := 0;
    IF recipeIn.recipeID <> 0 THEN
        FOR tmp_idx := 1 TO 10 DO
            IF recipe[tmp_idx].recipeID = recipeIn.recipeID THEN
                tmp_foundIdx := tmp_idx;
                EXIT;
            END_IF;
        END_FOR;
    END_IF;

    IF tmp_foundIdx = 0 THEN
        error := TRUE;
        status := 16#8001;
    ELSE
        recipeQueryResult := recipe[tmp_foundIdx];
    END_IF;
END_IF;

// Add operation (PUB003)
IF tmp_TrigAdd.Q THEN
    tmp_found := FALSE;
    tmp_emptyIdx := 0;

    FOR tmp_idx := 1 TO 10 DO
        IF recipe[tmp_idx].recipeID = recipeIn.recipeID THEN
            tmp_found := TRUE;
            EXIT;
        END_IF;
        IF recipe[tmp_idx].recipeID = 0 AND tmp_emptyIdx = 0 THEN
            tmp_emptyIdx := tmp_idx;
        END_IF;
    END_FOR;

    IF tmp_found THEN
        error := TRUE;
        status := 16#8002;
    ELSIF tmp_emptyIdx = 0 THEN
        error := TRUE;
        status := 16#8003;
    ELSE
        recipe[tmp_emptyIdx] := recipeIn;
        recipeAdded := TRUE;
    END_IF;
END_IF;

// Delete operation (PUB004)
IF tmp_TrigDelete.Q THEN
    tmp_foundIdx := 0;
    IF recipeIn.recipeID <> 0 THEN
        FOR tmp_idx := 1 TO 10 DO
            IF recipe[tmp_idx].recipeID = recipeIn.recipeID THEN
                tmp_foundIdx := tmp_idx;
                EXIT;
            END_IF;
        END_FOR;
    END_IF;

    IF tmp_foundIdx = 0 THEN
        error := TRUE;
        status := 16#8004;
    ELSE
        recipe[tmp_foundIdx].recipeID := 0;
        recipeDeleted := TRUE;
    END_IF;
END_IF;

// Modify operation (PUB005)
IF tmp_TrigModify.Q THEN
    tmp_foundIdx := 0;
    IF recipeIn.recipeID <> 0 THEN
        FOR tmp_idx := 1 TO 10 DO
            IF recipe[tmp_idx].recipeID = recipeIn.recipeID THEN
                tmp_foundIdx := tmp_idx;
                EXIT;
            END_IF;
        END_FOR;
    END_IF;

    IF tmp_foundIdx = 0 THEN
        error := TRUE;
        status := 16#8005;
    ELSE
        recipe[tmp_foundIdx] := recipeIn;
        recipeModified := TRUE;
    END_IF;
END_IF;

END_FUNCTION_BLOCK

(* ---- public-hard-03.raw_candidate_02.st ---- *)
(*
ENGINEERING_CONTRACT
- recipeAdded/Deleted/Modified: rising-edge pulse outputs, TRUE only on the scan where the corresponding request succeeds; no retention; reset next scan (PUB003/004/005).
- error: rising-edge pulse, TRUE only on the scan where an operation fails; no retention; reset next scan (PUB002-005).
- status: WORD code, 0 by default, nonzero only during a failed operation scan (PUB002-005).
- recipeQueryResult: zero-cleared at the start of every scan; holds the full recipe only during a successful query scan (PUB002).
- recipe database: persistent through IN_OUT; add uses smallest empty slot, duplicate check; delete sets recipeID to 0; modify replaces the whole struct (PUB003/004/005).
- Simultaneous requests are processed in the order query, add, delete, modify; unspecified by PUB002-005.
- recipeID 0 is treated as nonexistent for query/delete/modify and as duplicate for add because 0 marks an empty slot (PUB001).
*)
(* CONTRACT_RULES [] *)
TYPE ST_Recipe :
STRUCT
    recipeID : INT;
    ingredientType : INT;
    ingredientRatio : REAL;
    productionTemperature : REAL;
END_STRUCT
END_TYPE

FUNCTION_BLOCK FB_RecipeManagement
VAR_INPUT
    addRecipe : BOOL;
    deleteRecipe : BOOL;
    modifyRecipe : BOOL;
    queryRecipe : BOOL;
    recipeIn : ST_Recipe;
END_VAR

VAR_OUTPUT
    recipeAdded : BOOL;
    recipeDeleted : BOOL;
    recipeModified : BOOL;
    recipeQueryResult : ST_Recipe;
    error : BOOL;
    status : WORD;
END_VAR

VAR_IN_OUT
    recipe : ARRAY[1..10] OF ST_Recipe;
END_VAR

VAR
    tmp_TrigAdd : R_TRIG;
    tmp_TrigDelete : R_TRIG;
    tmp_TrigModify : R_TRIG;
    tmp_TrigQuery : R_TRIG;
    tmp_idx : INT;
    tmp_found : BOOL;
    tmp_foundIdx : INT;
    tmp_emptyIdx : INT;
END_VAR

// Evaluate rising edges once per scan.
tmp_TrigAdd(CLK := addRecipe);
tmp_TrigDelete(CLK := deleteRecipe);
tmp_TrigModify(CLK := modifyRecipe);
tmp_TrigQuery(CLK := queryRecipe);

// Default outputs for this scan.
recipeAdded := FALSE;
recipeDeleted := FALSE;
recipeModified := FALSE;
error := FALSE;
status := 0;

// Clear query result each scan; successful query will overwrite later.
recipeQueryResult.recipeID := 0;
recipeQueryResult.ingredientType := 0;
recipeQueryResult.ingredientRatio := 0.0;
recipeQueryResult.productionTemperature := 0.0;

// Query operation (PUB002)
IF tmp_TrigQuery.Q THEN
    tmp_foundIdx := 0;
    IF recipeIn.recipeID <> 0 THEN
        FOR tmp_idx := 1 TO 10 DO
            IF recipe[tmp_idx].recipeID = recipeIn.recipeID THEN
                tmp_foundIdx := tmp_idx;
                EXIT;
            END_IF;
        END_FOR;
    END_IF;

    IF tmp_foundIdx = 0 THEN
        error := TRUE;
        status := 16#8001;
    ELSE
        recipeQueryResult := recipe[tmp_foundIdx];
    END_IF;
END_IF;

// Add operation (PUB003)
IF tmp_TrigAdd.Q THEN
    tmp_found := FALSE;
    tmp_emptyIdx := 0;

    FOR tmp_idx := 1 TO 10 DO
        IF recipe[tmp_idx].recipeID = recipeIn.recipeID THEN
            tmp_found := TRUE;
            EXIT;
        END_IF;
        IF recipe[tmp_idx].recipeID = 0 AND tmp_emptyIdx = 0 THEN
            tmp_emptyIdx := tmp_idx;
        END_IF;
    END_FOR;

    IF tmp_found THEN
        error := TRUE;
        status := 16#8002;
    ELSIF tmp_emptyIdx = 0 THEN
        error := TRUE;
        status := 16#8003;
    ELSE
        recipe[tmp_emptyIdx] := recipeIn;
        recipeAdded := TRUE;
    END_IF;
END_IF;

// Delete operation (PUB004)
IF tmp_TrigDelete.Q THEN
    tmp_foundIdx := 0;
    IF recipeIn.recipeID <> 0 THEN
        FOR tmp_idx := 1 TO 10 DO
            IF recipe[tmp_idx].recipeID = recipeIn.recipeID THEN
                tmp_foundIdx := tmp_idx;
                EXIT;
            END_IF;
        END_FOR;
    END_IF;

    IF tmp_foundIdx = 0 THEN
        error := TRUE;
        status := 16#8004;
    ELSE
        recipe[tmp_foundIdx].recipeID := 0;
        recipeDeleted := TRUE;
    END_IF;
END_IF;

// Modify operation (PUB005)
IF tmp_TrigModify.Q THEN
    tmp_foundIdx := 0;
    IF recipeIn.recipeID <> 0 THEN
        FOR tmp_idx := 1 TO 10 DO
            IF recipe[tmp_idx].recipeID = recipeIn.recipeID THEN
                tmp_foundIdx := tmp_idx;
                EXIT;
            END_IF;
        END_FOR;
    END_IF;

    IF tmp_foundIdx = 0 THEN
        error := TRUE;
        status := 16#8005;
    ELSE
        recipe[tmp_foundIdx] := recipeIn;
        recipeModified := TRUE;
    END_IF;
END_IF;

END_FUNCTION_BLOCK

(* ---- public-hard-04.candidate_01.st ---- *)
(*
ENGINEERING_CONTRACT
1. elementCount: stored queue count; initial 0; reset->0; enqueue +1 on success;
   dequeue -1 on success; retained otherwise; range 0..capacity (PUB004).
2. status: per-scan combinational; default 16#0000 every invocation; set 16#8001 only
   for empty dequeue and 16#8002 only for full enqueue (PUB005). Reset clears to 0 (PUB003).
3. queue state head/tail/count initialized from buffer bounds on first call;
   capacity = UPPER_BOUND-LOWER_BOUND+1; empty first call (PUB006).
4. enqueue/dequeue edge-triggered via R_TRIG; one request per rising edge;
   reset TRUE consumes/ignores all edges and has priority (PUB001,PUB002,PUB003).
5. enqueue reads item and writes buffer[tail] only when count<capacity.
   dequeue writes item from buffer[head] only when count>0; rejected requests leave item and buffer unchanged (PUB005).
6. VARIANT buffer/output: direct indexed copy with matching element type;
   buffer bounds and association fixed per instance (PUB001,PUB006).
7. Simultaneous enqueue and dequeue is prohibited by caller (PUB002);
   implementation processes dequeue then enqueue if violated.
8. Units: elementCount elements; status WORD exact codes; buffer indices follow actual lower/upper bounds.
*)
(* CONTRACT_RULES [] *)
FUNCTION_BLOCK FB
VAR_INPUT
    enqueue : BOOL;
    dequeue : BOOL;
    reset : BOOL;
END_VAR
VAR_OUTPUT
    elementCount : DINT;
    status : WORD;
END_VAR
VAR_IN_OUT
    item : VARIANT;
    buffer : VARIANT;
END_VAR
VAR
    local_enq_edge : R_TRIG;
    local_deq_edge : R_TRIG;
    local_enq_req : BOOL;
    local_deq_req : BOOL;
    local_initialized : BOOL;
    local_lower : DINT;
    local_upper : DINT;
    local_capacity : DINT;
    local_head : DINT;
    local_tail : DINT;
    local_count : DINT;
END_VAR

IF NOT local_initialized THEN
    local_lower := LOWER_BOUND(buffer, 1);
    local_upper := UPPER_BOUND(buffer, 1);
    local_capacity := local_upper - local_lower + 1;
    IF local_capacity < 0 THEN
        local_capacity := 0;
    END_IF;
    local_head := local_lower;
    local_tail := local_lower;
    local_count := 0;
    local_initialized := TRUE;
END_IF;

elementCount := local_count;
status := WORD#16#0000;

local_enq_edge(CLK := enqueue);
local_deq_edge(CLK := dequeue);
local_enq_req := local_enq_edge.Q;
local_deq_req := local_deq_edge.Q;

IF reset THEN
    local_count := 0;
    local_head := local_lower;
    local_tail := local_lower;
    elementCount := 0;
    status := WORD#16#0000;
ELSE
    IF local_deq_req THEN
        IF local_count <= 0 THEN
            status := WORD#16#8001;
        ELSE
            item := buffer[local_head];
            local_head := local_head + 1;
            IF local_head > local_upper THEN
                local_head := local_lower;
            END_IF;
            local_count := local_count - 1;
            status := WORD#16#0000;
        END_IF;
    END_IF;

    IF local_enq_req THEN
        IF local_count >= local_capacity THEN
            status := WORD#16#8002;
        ELSE
            buffer[local_tail] := item;
            local_tail := local_tail + 1;
            IF local_tail > local_upper THEN
                local_tail := local_lower;
            END_IF;
            local_count := local_count + 1;
            status := WORD#16#0000;
        END_IF;
    END_IF;
END_IF;

elementCount := local_count;
END_FUNCTION_BLOCK

(* ---- public-hard-04.raw_candidate_01.st ---- *)
(*
ENGINEERING_CONTRACT
1. elementCount: stored queue count; initial 0; reset->0; enqueue +1 on success;
   dequeue -1 on success; retained otherwise; range 0..capacity (PUB004).
2. status: per-scan combinational; default 16#0000 every invocation; set 16#8001 only
   for empty dequeue and 16#8002 only for full enqueue (PUB005). Reset clears to 0 (PUB003).
3. queue state head/tail/count initialized from buffer bounds on first call;
   capacity = UPPER_BOUND-LOWER_BOUND+1; empty first call (PUB006).
4. enqueue/dequeue edge-triggered via R_TRIG; one request per rising edge;
   reset TRUE consumes/ignores all edges and has priority (PUB001,PUB002,PUB003).
5. enqueue reads item and writes buffer[tail] only when count<capacity.
   dequeue writes item from buffer[head] only when count>0; rejected requests leave item and buffer unchanged (PUB005).
6. VARIANT buffer/output: direct indexed copy with matching element type;
   buffer bounds and association fixed per instance (PUB001,PUB006).
7. Simultaneous enqueue and dequeue is prohibited by caller (PUB002);
   implementation processes dequeue then enqueue if violated.
8. Units: elementCount elements; status WORD exact codes; buffer indices follow actual lower/upper bounds.
*)
(* CONTRACT_RULES [] *)
FUNCTION_BLOCK FB
VAR_INPUT
    enqueue : BOOL;
    dequeue : BOOL;
    reset : BOOL;
END_VAR
VAR_OUTPUT
    elementCount : DINT;
    status : WORD;
END_VAR
VAR_IN_OUT
    item : VARIANT;
    buffer : VARIANT;
END_VAR
VAR
    local_enq_edge : R_TRIG;
    local_deq_edge : R_TRIG;
    local_enq_req : BOOL;
    local_deq_req : BOOL;
    local_initialized : BOOL;
    local_lower : DINT;
    local_upper : DINT;
    local_capacity : DINT;
    local_head : DINT;
    local_tail : DINT;
    local_count : DINT;
END_VAR

IF NOT local_initialized THEN
    local_lower := LOWER_BOUND(buffer, 1);
    local_upper := UPPER_BOUND(buffer, 1);
    local_capacity := local_upper - local_lower + 1;
    IF local_capacity < 0 THEN
        local_capacity := 0;
    END_IF;
    local_head := local_lower;
    local_tail := local_lower;
    local_count := 0;
    local_initialized := TRUE;
END_IF;

elementCount := local_count;
status := WORD#16#0000;

local_enq_edge(CLK := enqueue);
local_deq_edge(CLK := dequeue);
local_enq_req := local_enq_edge.Q;
local_deq_req := local_deq_edge.Q;

IF reset THEN
    local_count := 0;
    local_head := local_lower;
    local_tail := local_lower;
    elementCount := 0;
    status := WORD#16#0000;
ELSE
    IF local_deq_req THEN
        IF local_count <= 0 THEN
            status := WORD#16#8001;
        ELSE
            item := buffer[local_head];
            local_head := local_head + 1;
            IF local_head > local_upper THEN
                local_head := local_lower;
            END_IF;
            local_count := local_count - 1;
            status := WORD#16#0000;
        END_IF;
    END_IF;

    IF local_enq_req THEN
        IF local_count >= local_capacity THEN
            status := WORD#16#8002;
        ELSE
            buffer[local_tail] := item;
            local_tail := local_tail + 1;
            IF local_tail > local_upper THEN
                local_tail := local_lower;
            END_IF;
            local_count := local_count + 1;
            status := WORD#16#0000;
        END_IF;
    END_IF;
END_IF;

elementCount := local_count;
END_FUNCTION_BLOCK

(* ---- public-hard-05.candidate_01.st ---- *)
FUNCTION_BLOCK MechanicalArmControl
VAR_INPUT
    ManualMode : BOOL;
    SingleStepMode : BOOL;
    SingleCycleMode : BOOL;
    ContinuousMode : BOOL;
    EmergencyStop : BOOL;
    Start : BOOL;
    DownButton : BOOL;
    UpButton : BOOL;
    LeftButton : BOOL;
    RightButton : BOOL;
    GripButton : BOOL;
    ReleaseButton : BOOL;
    DownLimitSwitch : BOOL;
    UpLimitSwitch : BOOL;
    LeftLimitSwitch : BOOL;
    RightLimitSwitch : BOOL;
    GripLimitSwitch : BOOL;
    ReleaseLimitSwitch : BOOL;
END_VAR
VAR_OUTPUT
    MoveDown : BOOL;
    MoveUp : BOOL;
    MoveLeft : BOOL;
    MoveRight : BOOL;
    ActivateGrip : BOOL;
    ActivateRelease : BOOL;
END_VAR
VAR
    local_startR : R_TRIG;
    tmp_start_pulse : BOOL;
    tmp_not_estop : BOOL;
    tmp_ss_step : INT := 0;
    tmp_ss_busy : BOOL := FALSE;
    tmp_auto_running : BOOL := FALSE;
    tmp_auto_step : INT := 0;
    tmp_cmd_step : INT := 0;
    tmp_cmd_active : BOOL := FALSE;
    tmp_limit_reached : BOOL := FALSE;
END_VAR

(* ENGINEERING_CONTRACT
   Outputs MoveDown/Up/Left/Right/ActivateGrip/ActivateRelease:
   - Activate: manual while button=1, not at axis limit, and no opposite button (PUB001,PUB020); auto while current step active.
   - Retain: none latching; auto sequence state retained until completion/estop.
   - Reset: EmergencyStop=FALSE forces all outputs off and resets auto/single-step state (PUB005).
   - Same-scan: on limit true, previous output off; auto cycle can start next output in same scan (PUB003,PUB004).
   - Manual opposite-direction conflict inhibits both (PUB001 + shared rule).
   - Single-step Start edge only when not busy; ignored during running action (PUB002).
   - Single-cycle/continuous Start edge only when not running; continuous wraps at left completion (PUB003,PUB004).
   - Steps 0..7 = down, grip, up, right, down, release, up, left.
   - Grip/Release completion via GripLimitSwitch/ReleaseLimitSwitch (PUB001,PUB002).
   - Unspecified: mode change outside selected branch aborts/pauses per branch.
*)

(* CONTRACT_RULES [] *)

MoveDown := FALSE;
MoveUp := FALSE;
MoveLeft := FALSE;
MoveRight := FALSE;
ActivateGrip := FALSE;
ActivateRelease := FALSE;

tmp_not_estop := EmergencyStop; (* TRUE means no emergency stop triggered *)

local_startR(CLK := Start);
tmp_start_pulse := local_startR.Q;

tmp_cmd_active := FALSE;
tmp_cmd_step := 0;

IF NOT tmp_not_estop THEN
    tmp_ss_step := 0;
    tmp_ss_busy := FALSE;
    tmp_auto_running := FALSE;
    tmp_auto_step := 0;
    RETURN;
END_IF;

IF ManualMode THEN
    IF DownButton AND NOT UpButton AND NOT DownLimitSwitch THEN
        MoveDown := TRUE;
    END_IF;
    IF UpButton AND NOT DownButton AND NOT UpLimitSwitch THEN
        MoveUp := TRUE;
    END_IF;
    IF LeftButton AND NOT RightButton AND NOT LeftLimitSwitch THEN
        MoveLeft := TRUE;
    END_IF;
    IF RightButton AND NOT LeftButton AND NOT RightLimitSwitch THEN
        MoveRight := TRUE;
    END_IF;
    IF GripButton AND NOT ReleaseButton AND NOT GripLimitSwitch THEN
        ActivateGrip := TRUE;
    END_IF;
    IF ReleaseButton AND NOT GripButton AND NOT ReleaseLimitSwitch THEN
        ActivateRelease := TRUE;
    END_IF;

ELSIF SingleStepMode THEN
    IF tmp_start_pulse AND NOT tmp_ss_busy THEN
        tmp_ss_busy := TRUE;
    END_IF;

    IF tmp_ss_busy THEN
        tmp_limit_reached := FALSE;
        CASE tmp_ss_step OF
            0: tmp_limit_reached := DownLimitSwitch;
            1: tmp_limit_reached := GripLimitSwitch;
            2: tmp_limit_reached := UpLimitSwitch;
            3: tmp_limit_reached := RightLimitSwitch;
            4: tmp_limit_reached := DownLimitSwitch;
            5: tmp_limit_reached := ReleaseLimitSwitch;
            6: tmp_limit_reached := UpLimitSwitch;
            7: tmp_limit_reached := LeftLimitSwitch;
        END_CASE;

        IF tmp_limit_reached THEN
            tmp_ss_busy := FALSE;
            tmp_ss_step := tmp_ss_step + 1;
            IF tmp_ss_step > 7 THEN
                tmp_ss_step := 0;
            END_IF;
        ELSE
            tmp_cmd_step := tmp_ss_step;
            tmp_cmd_active := TRUE;
        END_IF;
    END_IF;

ELSIF SingleCycleMode OR ContinuousMode THEN
    IF tmp_start_pulse AND NOT tmp_auto_running THEN
        tmp_auto_running := TRUE;
        tmp_auto_step := 0;
    END_IF;

    IF tmp_auto_running THEN
        tmp_limit_reached := FALSE;
        CASE tmp_auto_step OF
            0: tmp_limit_reached := DownLimitSwitch;
            1: tmp_limit_reached := GripLimitSwitch;
            2: tmp_limit_reached := UpLimitSwitch;
            3: tmp_limit_reached := RightLimitSwitch;
            4: tmp_limit_reached := DownLimitSwitch;
            5: tmp_limit_reached := ReleaseLimitSwitch;
            6: tmp_limit_reached := UpLimitSwitch;
            7: tmp_limit_reached := LeftLimitSwitch;
        END_CASE;

        IF tmp_limit_reached THEN
            IF tmp_auto_step = 7 THEN
                IF ContinuousMode THEN
                    tmp_auto_step := 0; (* start next cycle *)
                ELSE
                    tmp_auto_running := FALSE;
                    tmp_auto_step := 0;
                END_IF;
            ELSE
                tmp_auto_step := tmp_auto_step + 1;
            END_IF;
        END_IF;

        IF tmp_auto_running THEN
            tmp_cmd_step := tmp_auto_step;
            tmp_cmd_active := TRUE;
        END_IF;
    END_IF;
END_IF;

IF tmp_cmd_active THEN
    CASE tmp_cmd_step OF
        0: MoveDown := TRUE;
        1: ActivateGrip := TRUE;
        2: MoveUp := TRUE;
        3: MoveRight := TRUE;
        4: MoveDown := TRUE;
        5: ActivateRelease := TRUE;
        6: MoveUp := TRUE;
        7: MoveLeft := TRUE;
    END_CASE;
END_IF;

END_FUNCTION_BLOCK

(* ---- public-hard-05.candidate_02.st ---- *)
FUNCTION_BLOCK MechanicalArmControl
VAR_INPUT
    ManualMode : BOOL;
    SingleStepMode : BOOL;
    SingleCycleMode : BOOL;
    ContinuousMode : BOOL;
    EmergencyStop : BOOL;
    Start : BOOL;
    DownButton : BOOL;
    UpButton : BOOL;
    LeftButton : BOOL;
    RightButton : BOOL;
    GripButton : BOOL;
    ReleaseButton : BOOL;
    DownLimitSwitch : BOOL;
    UpLimitSwitch : BOOL;
    LeftLimitSwitch : BOOL;
    RightLimitSwitch : BOOL;
    GripLimitSwitch : BOOL;
    ReleaseLimitSwitch : BOOL;
END_VAR
VAR_OUTPUT
    MoveDown : BOOL;
    MoveUp : BOOL;
    MoveLeft : BOOL;
    MoveRight : BOOL;
    ActivateGrip : BOOL;
    ActivateRelease : BOOL;
END_VAR
VAR
    local_startR : R_TRIG;
    tmp_first_scan : BOOL := TRUE;
    tmp_start_pulse : BOOL;
    tmp_not_estop : BOOL;
    tmp_ss_step : INT := 0;
    tmp_ss_busy : BOOL := FALSE;
    tmp_auto_running : BOOL := FALSE;
    tmp_auto_step : INT := 0;
    tmp_cmd_step : INT := 0;
    tmp_cmd_active : BOOL := FALSE;
    tmp_limit_reached : BOOL := FALSE;
END_VAR

(* ENGINEERING_CONTRACT
   Outputs MoveDown/Up/Left/Right/ActivateGrip/ActivateRelease:
   - Activate: manual while button=1, not at axis limit, and no opposite button (PUB001,PUB020); auto while current step active.
   - Retain: none latching; auto sequence state retained until completion/estop.
   - Reset: EmergencyStop=FALSE forces all outputs off and resets auto/single-step state (PUB005).
   - Same-scan: on limit true, previous output off; auto cycle can start next output in same scan (PUB003,PUB004).
   - Manual opposite-direction conflict inhibits both (PUB001 + shared rule).
   - Single-step Start edge only when not busy; ignored during running action (PUB002).
   - Single-cycle/continuous Start edge only when not running; continuous wraps at left completion (PUB003,PUB004).
   - Steps 0..7 = down, grip, up, right, down, release, up, left.
   - Grip/Release completion via GripLimitSwitch/ReleaseLimitSwitch (PUB001,PUB002).
   - Unspecified: mode change outside selected branch aborts/pauses per branch.
*)

(* CONTRACT_RULES [] *)

MoveDown := FALSE;
MoveUp := FALSE;
MoveLeft := FALSE;
MoveRight := FALSE;
ActivateGrip := FALSE;
ActivateRelease := FALSE;

tmp_not_estop := EmergencyStop; (* TRUE means no emergency stop triggered *)

local_startR(CLK := Start);
tmp_start_pulse := local_startR.Q AND NOT tmp_first_scan;
tmp_first_scan := FALSE;

tmp_cmd_active := FALSE;
tmp_cmd_step := 0;

IF NOT tmp_not_estop THEN
    tmp_ss_step := 0;
    tmp_ss_busy := FALSE;
    tmp_auto_running := FALSE;
    tmp_auto_step := 0;
    RETURN;
END_IF;

IF ManualMode THEN
    IF DownButton AND NOT UpButton AND NOT DownLimitSwitch THEN
        MoveDown := TRUE;
    END_IF;
    IF UpButton AND NOT DownButton AND NOT UpLimitSwitch THEN
        MoveUp := TRUE;
    END_IF;
    IF LeftButton AND NOT RightButton AND NOT LeftLimitSwitch THEN
        MoveLeft := TRUE;
    END_IF;
    IF RightButton AND NOT LeftButton AND NOT RightLimitSwitch THEN
        MoveRight := TRUE;
    END_IF;
    IF GripButton AND NOT ReleaseButton AND NOT GripLimitSwitch THEN
        ActivateGrip := TRUE;
    END_IF;
    IF ReleaseButton AND NOT GripButton AND NOT ReleaseLimitSwitch THEN
        ActivateRelease := TRUE;
    END_IF;

ELSIF SingleStepMode THEN
    IF tmp_start_pulse AND NOT tmp_ss_busy THEN
        tmp_ss_busy := TRUE;
    END_IF;

    IF tmp_ss_busy THEN
        tmp_limit_reached := FALSE;
        CASE tmp_ss_step OF
            0: tmp_limit_reached := DownLimitSwitch;
            1: tmp_limit_reached := GripLimitSwitch;
            2: tmp_limit_reached := UpLimitSwitch;
            3: tmp_limit_reached := RightLimitSwitch;
            4: tmp_limit_reached := DownLimitSwitch;
            5: tmp_limit_reached := ReleaseLimitSwitch;
            6: tmp_limit_reached := UpLimitSwitch;
            7: tmp_limit_reached := LeftLimitSwitch;
        END_CASE;

        IF tmp_limit_reached THEN
            tmp_ss_busy := FALSE;
            tmp_ss_step := tmp_ss_step + 1;
            IF tmp_ss_step > 7 THEN
                tmp_ss_step := 0;
            END_IF;
        ELSE
            tmp_cmd_step := tmp_ss_step;
            tmp_cmd_active := TRUE;
        END_IF;
    END_IF;

ELSIF SingleCycleMode OR ContinuousMode THEN
    IF tmp_start_pulse AND NOT tmp_auto_running THEN
        tmp_auto_running := TRUE;
        tmp_auto_step := 0;
    END_IF;

    IF tmp_auto_running THEN
        tmp_limit_reached := FALSE;
        CASE tmp_auto_step OF
            0: tmp_limit_reached := DownLimitSwitch;
            1: tmp_limit_reached := GripLimitSwitch;
            2: tmp_limit_reached := UpLimitSwitch;
            3: tmp_limit_reached := RightLimitSwitch;
            4: tmp_limit_reached := DownLimitSwitch;
            5: tmp_limit_reached := ReleaseLimitSwitch;
            6: tmp_limit_reached := UpLimitSwitch;
            7: tmp_limit_reached := LeftLimitSwitch;
        END_CASE;

        IF tmp_limit_reached THEN
            IF tmp_auto_step = 7 THEN
                IF ContinuousMode THEN
                    tmp_auto_step := 0; (* start next cycle *)
                ELSE
                    tmp_auto_running := FALSE;
                    tmp_auto_step := 0;
                END_IF;
            ELSE
                tmp_auto_step := tmp_auto_step + 1;
            END_IF;
        END_IF;

        IF tmp_auto_running THEN
            tmp_cmd_step := tmp_auto_step;
            tmp_cmd_active := TRUE;
        END_IF;
    END_IF;
END_IF;

IF tmp_cmd_active THEN
    CASE tmp_cmd_step OF
        0: MoveDown := TRUE;
        1: ActivateGrip := TRUE;
        2: MoveUp := TRUE;
        3: MoveRight := TRUE;
        4: MoveDown := TRUE;
        5: ActivateRelease := TRUE;
        6: MoveUp := TRUE;
        7: MoveLeft := TRUE;
    END_CASE;
END_IF;

END_FUNCTION_BLOCK

(* ---- public-hard-05.candidate_03.st ---- *)
FUNCTION_BLOCK MechanicalArmControl
VAR_INPUT
    ManualMode : BOOL;
    SingleStepMode : BOOL;
    SingleCycleMode : BOOL;
    ContinuousMode : BOOL;
    EmergencyStop : BOOL;
    Start : BOOL;
    DownButton : BOOL;
    UpButton : BOOL;
    LeftButton : BOOL;
    RightButton : BOOL;
    GripButton : BOOL;
    ReleaseButton : BOOL;
    DownLimitSwitch : BOOL;
    UpLimitSwitch : BOOL;
    LeftLimitSwitch : BOOL;
    RightLimitSwitch : BOOL;
    GripLimitSwitch : BOOL;
    ReleaseLimitSwitch : BOOL;
END_VAR
VAR_OUTPUT
    MoveDown : BOOL;
    MoveUp : BOOL;
    MoveLeft : BOOL;
    MoveRight : BOOL;
    ActivateGrip : BOOL;
    ActivateRelease : BOOL;
END_VAR
VAR
    local_startR : R_TRIG;
    tmp_start_pulse : BOOL;
    tmp_not_estop : BOOL;
    tmp_ss_step : INT := 0;
    tmp_ss_busy : BOOL := FALSE;
    tmp_auto_running : BOOL := FALSE;
    tmp_auto_step : INT := 0;
    tmp_cmd_step : INT := 0;
    tmp_cmd_active : BOOL := FALSE;
    tmp_limit_reached : BOOL := FALSE;
END_VAR

(* ENGINEERING_CONTRACT
   Outputs MoveDown/Up/Left/Right/ActivateGrip/ActivateRelease:
   - Activate: manual while button=1, not at axis limit, and no opposite button (PUB001,PUB020); auto while current step active.
   - Retain: none latching; auto sequence state retained until completion/estop.
   - Reset: EmergencyStop=FALSE forces all outputs off and resets auto/single-step state (PUB005).
   - Same-scan: on limit true, previous output off; auto cycle can start next output in same scan (PUB003,PUB004).
   - Manual opposite-direction conflict inhibits both (PUB001 + shared rule).
   - Single-step Start edge only when not busy; ignored during running action (PUB002).
   - Single-cycle/continuous Start edge only when not running; continuous wraps at left completion (PUB003,PUB004).
   - Steps 0..7 = down, grip, up, right, down, release, up, left.
   - Grip/Release completion via GripLimitSwitch/ReleaseLimitSwitch (PUB001,PUB002).
   - Unspecified: mode change outside selected branch aborts/pauses per branch.
*)

(* CONTRACT_RULES [] *)

MoveDown := FALSE;
MoveUp := FALSE;
MoveLeft := FALSE;
MoveRight := FALSE;
ActivateGrip := FALSE;
ActivateRelease := FALSE;

tmp_not_estop := EmergencyStop; (* TRUE means no emergency stop triggered *)

local_startR(CLK := Start);
tmp_start_pulse := local_startR.Q;

tmp_cmd_active := FALSE;
tmp_cmd_step := 0;

IF NOT tmp_not_estop THEN
    tmp_ss_step := 0;
    tmp_ss_busy := FALSE;
    tmp_auto_running := FALSE;
    tmp_auto_step := 0;
    RETURN;
END_IF;

IF ManualMode THEN
    IF DownButton AND NOT UpButton AND NOT DownLimitSwitch THEN
        MoveDown := TRUE;
    END_IF;
    IF UpButton AND NOT DownButton AND NOT UpLimitSwitch THEN
        MoveUp := TRUE;
    END_IF;
    IF LeftButton AND NOT RightButton AND NOT LeftLimitSwitch THEN
        MoveLeft := TRUE;
    END_IF;
    IF RightButton AND NOT LeftButton AND NOT RightLimitSwitch THEN
        MoveRight := TRUE;
    END_IF;
    IF GripButton AND NOT ReleaseButton AND NOT GripLimitSwitch THEN
        ActivateGrip := TRUE;
    END_IF;
    IF ReleaseButton AND NOT GripButton AND NOT ReleaseLimitSwitch THEN
        ActivateRelease := TRUE;
    END_IF;

ELSIF SingleStepMode THEN
    IF tmp_start_pulse AND NOT tmp_ss_busy THEN
        tmp_ss_busy := TRUE;
    END_IF;

    IF tmp_ss_busy THEN
        tmp_limit_reached := FALSE;
        CASE tmp_ss_step OF
            0: tmp_limit_reached := DownLimitSwitch;
            1: tmp_limit_reached := GripLimitSwitch;
            2: tmp_limit_reached := UpLimitSwitch;
            3: tmp_limit_reached := RightLimitSwitch;
            4: tmp_limit_reached := DownLimitSwitch;
            5: tmp_limit_reached := ReleaseLimitSwitch;
            6: tmp_limit_reached := UpLimitSwitch;
            7: tmp_limit_reached := LeftLimitSwitch;
        END_CASE;

        IF tmp_limit_reached THEN
            tmp_ss_busy := FALSE;
            tmp_ss_step := tmp_ss_step + 1;
            IF tmp_ss_step > 7 THEN
                tmp_ss_step := 0;
            END_IF;
        ELSE
            tmp_cmd_step := tmp_ss_step;
            tmp_cmd_active := TRUE;
        END_IF;
    END_IF;

ELSIF SingleCycleMode OR ContinuousMode THEN
    IF tmp_start_pulse AND NOT tmp_auto_running THEN
        tmp_auto_running := TRUE;
        tmp_auto_step := 0;
    END_IF;

    IF tmp_auto_running THEN
        tmp_limit_reached := FALSE;
        CASE tmp_auto_step OF
            0: tmp_limit_reached := DownLimitSwitch;
            1: tmp_limit_reached := GripLimitSwitch;
            2: tmp_limit_reached := UpLimitSwitch;
            3: tmp_limit_reached := RightLimitSwitch;
            4: tmp_limit_reached := DownLimitSwitch;
            5: tmp_limit_reached := ReleaseLimitSwitch;
            6: tmp_limit_reached := UpLimitSwitch;
            7: tmp_limit_reached := LeftLimitSwitch;
        END_CASE;

        IF tmp_limit_reached THEN
            IF tmp_auto_step = 7 THEN
                IF ContinuousMode THEN
                    tmp_auto_step := 0; (* start next cycle *)
                ELSE
                    tmp_auto_running := FALSE;
                    tmp_auto_step := 0;
                END_IF;
            ELSE
                tmp_auto_step := tmp_auto_step + 1;
            END_IF;
        END_IF;

        IF tmp_auto_running THEN
            tmp_cmd_step := tmp_auto_step;
            tmp_cmd_active := TRUE;
        END_IF;
    END_IF;
END_IF;

IF tmp_cmd_active THEN
    CASE tmp_cmd_step OF
        0: MoveDown := TRUE;
        1: ActivateGrip := TRUE;
        2: MoveUp := TRUE;
        3: MoveRight := TRUE;
        4: MoveDown := TRUE;
        5: ActivateRelease := TRUE;
        6: MoveUp := TRUE;
        7: MoveLeft := TRUE;
    END_CASE;
END_IF;

END_FUNCTION_BLOCK

(* ---- public-hard-05.patch_base_02.st ---- *)
FUNCTION_BLOCK MechanicalArmControl
VAR_INPUT
    ManualMode : BOOL;
    SingleStepMode : BOOL;
    SingleCycleMode : BOOL;
    ContinuousMode : BOOL;
    EmergencyStop : BOOL;
    Start : BOOL;
    DownButton : BOOL;
    UpButton : BOOL;
    LeftButton : BOOL;
    RightButton : BOOL;
    GripButton : BOOL;
    ReleaseButton : BOOL;
    DownLimitSwitch : BOOL;
    UpLimitSwitch : BOOL;
    LeftLimitSwitch : BOOL;
    RightLimitSwitch : BOOL;
    GripLimitSwitch : BOOL;
    ReleaseLimitSwitch : BOOL;
END_VAR
VAR_OUTPUT
    MoveDown : BOOL;
    MoveUp : BOOL;
    MoveLeft : BOOL;
    MoveRight : BOOL;
    ActivateGrip : BOOL;
    ActivateRelease : BOOL;
END_VAR
VAR
    local_startR : R_TRIG;
    tmp_start_pulse : BOOL;
    tmp_not_estop : BOOL;
    tmp_ss_step : INT := 0;
    tmp_ss_busy : BOOL := FALSE;
    tmp_auto_running : BOOL := FALSE;
    tmp_auto_step : INT := 0;
    tmp_cmd_step : INT := 0;
    tmp_cmd_active : BOOL := FALSE;
    tmp_limit_reached : BOOL := FALSE;
END_VAR

(* ENGINEERING_CONTRACT
   Outputs MoveDown/Up/Left/Right/ActivateGrip/ActivateRelease:
   - Activate: manual while button=1, not at axis limit, and no opposite button (PUB001,PUB020); auto while current step active.
   - Retain: none latching; auto sequence state retained until completion/estop.
   - Reset: EmergencyStop=FALSE forces all outputs off and resets auto/single-step state (PUB005).
   - Same-scan: on limit true, previous output off; auto cycle can start next output in same scan (PUB003,PUB004).
   - Manual opposite-direction conflict inhibits both (PUB001 + shared rule).
   - Single-step Start edge only when not busy; ignored during running action (PUB002).
   - Single-cycle/continuous Start edge only when not running; continuous wraps at left completion (PUB003,PUB004).
   - Steps 0..7 = down, grip, up, right, down, release, up, left.
   - Grip/Release completion via GripLimitSwitch/ReleaseLimitSwitch (PUB001,PUB002).
   - Unspecified: mode change outside selected branch aborts/pauses per branch.
*)

(* CONTRACT_RULES [] *)

MoveDown := FALSE;
MoveUp := FALSE;
MoveLeft := FALSE;
MoveRight := FALSE;
ActivateGrip := FALSE;
ActivateRelease := FALSE;

tmp_not_estop := EmergencyStop; (* TRUE means no emergency stop triggered *)

local_startR(CLK := Start);
tmp_start_pulse := local_startR.Q;

tmp_cmd_active := FALSE;
tmp_cmd_step := 0;

IF NOT tmp_not_estop THEN
    tmp_ss_step := 0;
    tmp_ss_busy := FALSE;
    tmp_auto_running := FALSE;
    tmp_auto_step := 0;
    RETURN;
END_IF;

IF ManualMode THEN
    IF DownButton AND NOT UpButton AND NOT DownLimitSwitch THEN
        MoveDown := TRUE;
    END_IF;
    IF UpButton AND NOT DownButton AND NOT UpLimitSwitch THEN
        MoveUp := TRUE;
    END_IF;
    IF LeftButton AND NOT RightButton AND NOT LeftLimitSwitch THEN
        MoveLeft := TRUE;
    END_IF;
    IF RightButton AND NOT LeftButton AND NOT RightLimitSwitch THEN
        MoveRight := TRUE;
    END_IF;
    IF GripButton AND NOT ReleaseButton AND NOT GripLimitSwitch THEN
        ActivateGrip := TRUE;
    END_IF;
    IF ReleaseButton AND NOT GripButton AND NOT ReleaseLimitSwitch THEN
        ActivateRelease := TRUE;
    END_IF;

ELSIF SingleStepMode THEN
    IF tmp_start_pulse AND NOT tmp_ss_busy THEN
        tmp_ss_busy := TRUE;
    END_IF;

    IF tmp_ss_busy THEN
        tmp_limit_reached := FALSE;
        CASE tmp_ss_step OF
            0: tmp_limit_reached := DownLimitSwitch;
            1: tmp_limit_reached := GripLimitSwitch;
            2: tmp_limit_reached := UpLimitSwitch;
            3: tmp_limit_reached := RightLimitSwitch;
            4: tmp_limit_reached := DownLimitSwitch;
            5: tmp_limit_reached := ReleaseLimitSwitch;
            6: tmp_limit_reached := UpLimitSwitch;
            7: tmp_limit_reached := LeftLimitSwitch;
        END_CASE;

        IF tmp_limit_reached THEN
            tmp_ss_busy := FALSE;
            tmp_ss_step := tmp_ss_step + 1;
            IF tmp_ss_step > 7 THEN
                tmp_ss_step := 0;
            END_IF;
        ELSE
            tmp_cmd_step := tmp_ss_step;
            tmp_cmd_active := TRUE;
        END_IF;
    END_IF;

ELSIF SingleCycleMode OR ContinuousMode THEN
    IF tmp_start_pulse AND NOT tmp_auto_running THEN
        tmp_auto_running := TRUE;
        tmp_auto_step := 0;
    END_IF;

    IF tmp_auto_running THEN
        tmp_limit_reached := FALSE;
        CASE tmp_auto_step OF
            0: tmp_limit_reached := DownLimitSwitch;
            1: tmp_limit_reached := GripLimitSwitch;
            2: tmp_limit_reached := UpLimitSwitch;
            3: tmp_limit_reached := RightLimitSwitch;
            4: tmp_limit_reached := DownLimitSwitch;
            5: tmp_limit_reached := ReleaseLimitSwitch;
            6: tmp_limit_reached := UpLimitSwitch;
            7: tmp_limit_reached := LeftLimitSwitch;
        END_CASE;

        IF tmp_limit_reached THEN
            IF tmp_auto_step = 7 THEN
                IF ContinuousMode THEN
                    tmp_auto_step := 0; (* start next cycle *)
                ELSE
                    tmp_auto_running := FALSE;
                    tmp_auto_step := 0;
                END_IF;
            ELSE
                tmp_auto_step := tmp_auto_step + 1;
            END_IF;
        END_IF;

        IF tmp_auto_running THEN
            tmp_cmd_step := tmp_auto_step;
            tmp_cmd_active := TRUE;
        END_IF;
    END_IF;
END_IF;

IF tmp_cmd_active THEN
    CASE tmp_cmd_step OF
        0: MoveDown := TRUE;
        1: ActivateGrip := TRUE;
        2: MoveUp := TRUE;
        3: MoveRight := TRUE;
        4: MoveDown := TRUE;
        5: ActivateRelease := TRUE;
        6: MoveUp := TRUE;
        7: MoveLeft := TRUE;
    END_CASE;
END_IF;

END_FUNCTION_BLOCK
